(* IEC 61131-3 sources: rusty/tests/lit/cfc/blocks/function_chain, 2 files *)

(* ---- main.st ---- *)
FUNCTION main : DINT
    function_chain.seed := 3;
    function_chain.k := 4;
    function_chain();
    // chain: (seed + k) then (+ k) => (3 + 4) + 4
    // CHECK: result = 11
    printf('result = %d$N', function_chain.result);
END_FUNCTION

(* ---- myAdd.st ---- *)
FUNCTION myAdd : INT
    VAR_INPUT
        in1, in2: DINT;
    END_VAR

    VAR_OUTPUT
        myAddDoubled: DINT;
    END_VAR

    myAdd := in1 + in2;
    myAddDoubled := (in1 + in2) * 2;
END_FUNCTION
